Fanuc KAREL source: KT00876.KL

PROGRAM KT00876
%NOLOCKGROUP
VAR
  B1: BOOLEAN
  B2: BOOLEAN
  OUT: INTEGER
BEGIN
  B1 = TRUE
  B2 = FALSE
  B1 = TRUE
  B2 = FALSE
  OUT = TRUNC(B1)
END KT00876
